(* IEC 61131-3 sources: ATCMcontrol_Engineering/src/TargetBase/Libs/ATCM_IEC1131_3/table_25, 4 files *)

(* ---- ROL.st ---- *)
FUNCTION ROL : any_bit
VAR_INPUT
    IN : any_bit;
    N  : any_int;
END_VAR

(* we do not support DINT as second param *)
(*
overload bool(bool,dint)
inline
{
    %1
    %2
    dint_to_int
    rol_bool
}
overload byte(byte,dint)
inline
{
    %1
    %2
    dint_to_int
    rol_byte
}
overload word(word,dint)
inline
{
    %1
    %2
    dint_to_int
    rol_word
}
overload dword(dword,dint)
inline
{
    %1
    %2
    dint_to_int
    rol_dword
}
*)

overload bool(bool,int)   inline{ VMOP(rol_bool) }
overload byte(byte,int)   inline{ VMOP(rol_byte) }
overload word(word,int)   inline{ VMOP(rol_word) }
overload dword(dword,int) inline{ VMOP(rol_dword) }

(*
overload LWORD(LWORD,INT) inline{}
overload LWORD(LWORD,DINT) inline{}
*)
END_FUNCTION

(* ---- ROR.st ---- *)
FUNCTION ROR : any_bit
VAR_INPUT
    IN : any_bit;
    N  : any_int;
END_VAR

(* we do not support DINT as second param *)
(*
overload bool(bool,dint)
inline
{
    %1
    %2
    dint_to_int
    ror_bool
}
overload byte(byte,dint)
inline
{
    %1
    %2
    dint_to_int
    ror_byte
}
overload word(word,dint)
inline
{
    %1
    %2
    dint_to_int
    ror_word
}
overload dword(dword,dint)
inline
{
    %1
    %2
    dint_to_int
    ror_dword
}
*)

overload bool(bool,int)   inline{ VMOP(ror_bool) }
overload byte(byte,int)   inline{ VMOP(ror_byte) }
overload word(word,int)   inline{ VMOP(ror_word) }
overload dword(dword,int) inline{ VMOP(ror_dword) }

(*
overload LWORD(LWORD,INT) inline{}
overload LWORD(LWORD,DINT) inline{}
*)
END_FUNCTION

(* ---- SHL.st ---- *)
FUNCTION SHL : any_bit
VAR_INPUT
    IN : any_bit;
    N  : any_int;
END_VAR

(* we do not support DINT as second param *)
(*
overload bool(bool,dint)
inline
{
    %1
    %2
    dint_to_int
    shl_bool
}
overload byte(byte,dint)
inline
{
    %1
    %2
    dint_to_int
    shl_byte
}
overload word(word,dint)
inline
{
    %1
    %2
    dint_to_int
    shl_word
}
overload dword(dword,dint)
inline
{
    %1
    %2
    dint_to_int
    shl_dword
}
*)

overload bool(bool,int)   inline{ VMOP(shl_bool) }
overload byte(byte,int)   inline{ VMOP(shl_byte) }
overload word(word,int)   inline{ VMOP(shl_word) }
overload dword(dword,int) inline{ VMOP(shl_dword) }

(*
overload LWORD(LWORD,INT) inline{}
overload LWORD(LWORD,DINT) inline{}
*)
END_FUNCTION

(* ---- SHR.st ---- *)
FUNCTION SHR : any_bit
VAR_INPUT
    IN : any_bit;
    N  : any_int;
END_VAR

(* we do not support DINT as second param *)
(*
overload bool(bool,dint)
inline
{
    %1
    %2
    dint_to_int
    shr_bool
}
overload byte(byte,dint)
inline
{
    %1
    %2
    dint_to_int
    shr_byte
}
overload word(word,dint)
inline
{
    %1
    %2
    dint_to_int
    shr_word
}
overload dword(dword,dint)
inline
{
    %1
    %2
    dint_to_int
    shr_dword
}
*)

overload bool(bool,int)   inline{ VMOP(shr_bool) }
overload byte(byte,int)   inline{ VMOP(shr_byte) }
overload word(word,int)   inline{ VMOP(shr_word) }
overload dword(dword,int) inline{ VMOP(shr_dword) }

(*
overload LWORD(LWORD,INT) inline{}
overload LWORD(LWORD,DINT) inline{}
*)

END_FUNCTION
